(* PLC project p3_sfc_clean, Anonymous Benchmark Suite 1.0 *)
(* stored: creationDateTime 2026-08-25T00:00:00 *)

PROGRAM drive
  VAR_INPUT
    fwd : BOOL;
    rev : BOOL;
    maint : BOOL;
  END_VAR
  VAR_OUTPUT
    Motor_A : BOOL;
    Motor_B : BOOL;
  END_VAR

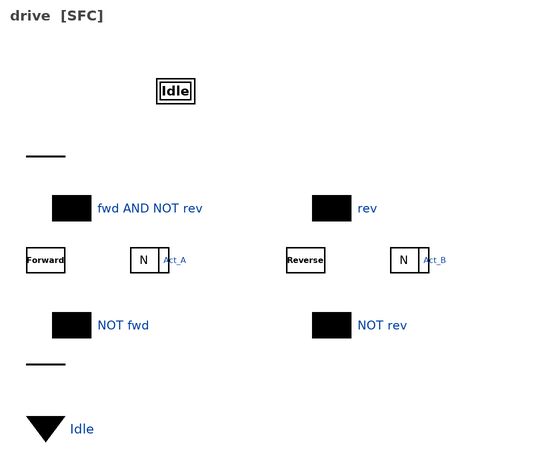
INITIAL_STEP Idle:
END_STEP
TRANSITION FROM Idle TO Forward
  := fwd AND NOT rev;
END_TRANSITION
TRANSITION FROM Idle TO Reverse
  := rev;
END_TRANSITION
STEP Forward:
  Act_A(N);
END_STEP
TRANSITION FROM Forward TO Idle
  := NOT fwd;
END_TRANSITION
STEP Reverse:
  Act_B(N);
END_STEP
TRANSITION FROM Reverse TO Idle
  := NOT rev;
END_TRANSITION

ACTION Act_A:
Motor_A := TRUE;
END_ACTION

ACTION Act_B:
Motor_B := TRUE;
END_ACTION

ACTION Act_Both:
Motor_A := TRUE;
Motor_B := TRUE;
END_ACTION
END_PROGRAM

CONFIGURATION Config0
  RESOURCE Res0 ON PLC
    TASK tcyclic(INTERVAL := T#10ms, PRIORITY := 0);
    PROGRAM inst0 WITH tcyclic : drive;
  END_RESOURCE
END_CONFIGURATION
